{attribute 'qualified_only'}
{attribute 'strict'}
{attribute 'to_string'}
TYPE E_OperationState :
(
    Idle  := 0,     // never started
    Busy  := 1,
    Done  := 2,
    Error := 3
);
END_TYPE

(* stored: Version 1.1.0.1
   DUT E_OperationState: Id {02c5dc91-cbd4-425e-92f8-3c0885740113} *)
